Fanuc KAREL source: KT00700.KL

PROGRAM KT00700
%NOLOCKGROUP
VAR
  C1: CONFIG
  C2: CONFIG
  OUT: INTEGER
BEGIN
  C1.CFG_FLIP = TRUE
  C2.CFG_FLIP = FALSE
  C1.CFG_FLIP = TRUE
  C2.CFG_FLIP = FALSE
  OUT = + C1
END KT00700
